Fanuc KAREL source: KB00022.KL

PROGRAM KB00022
%NOLOCKGROUP
%ENVIRONMENT MULTI
VAR
  P1: INTEGER
BEGIN
  P1 = 1
  CLEAR_SEMA(P1)
END KB00022
